(* IEC 61131-3 sources: plcassist-cli/packages/volt-lsp-iec/test-corpus/lenze-mid/Device/Plc Logic/Application/Library Manager/CAA Behaviour Model, 12 files *)

(* ---- VERSIONCONSTANTS.gvl ---- *)
VAR_GLOBAL
	GC_BYVERSION : BYTE := 1;
	GC_BYVERSION_1 : BYTE := 0;
END_VAR

(* ---- IFBCOMMAND.itf ---- *)
INTERFACE IFBCOMMAND
END_INTERFACE

METHOD PRVABORT : BOOL
END_METHOD

METHOD PRVCYCLICACTION : BOOL
END_METHOD

METHOD PRVRESETOUTPUTS : BOOL
END_METHOD

METHOD PRVSTART : BOOL
END_METHOD

(* ---- GETSUPPLIERVERSION.fun ---- *)
FUNCTION GETSUPPLIERVERSION : WORD
VAR_INPUT
	XDUMMY : BOOL;
END_VAR
END_FUNCTION

(* ---- ETRIG.fb ---- *)
FUNCTION_BLOCK ETRIG
VAR_INPUT
	XEXECUTE : BOOL;
END_VAR
VAR_OUTPUT
	XDONE : BOOL;
	XBUSY : BOOL;
	XERROR : BOOL;
END_VAR
VAR
	XPREVIOUSEXECUTE : BOOL;
	XPREVIOUSABORTINPROGRESS : BOOL;
	XABORTINPROGRESS : BOOL;
	IERROR : INT;
END_VAR
END_FUNCTION_BLOCK

METHOD PRVABORT : BOOL
END_METHOD

METHOD PRVCYCLICACTION : BOOL
END_METHOD

METHOD PRVRESETOUTPUTS : BOOL
END_METHOD

METHOD PRVSTART : BOOL
END_METHOD

(* ---- ETRIGA.fb ---- *)
FUNCTION_BLOCK ETRIGA
VAR_INPUT
	XEXECUTE : BOOL;
	XABORT : BOOL;
END_VAR
VAR_OUTPUT
	XDONE : BOOL;
	XBUSY : BOOL;
	XERROR : BOOL;
	XABORTED : BOOL;
END_VAR
VAR
	XPREVIOUSABORTINPROGRESS : BOOL;
	XPREVIOUSEXECUTE : BOOL;
	XABORTINPROGRESS : BOOL;
	IERROR : INT;
END_VAR
END_FUNCTION_BLOCK

METHOD PRVABORT : BOOL
END_METHOD

METHOD PRVCYCLICACTION : BOOL
END_METHOD

METHOD PRVRESETOUTPUTS : BOOL
END_METHOD

METHOD PRVSTART : BOOL
END_METHOD

(* ---- ETRIGTL.fb ---- *)
FUNCTION_BLOCK ETRIGTL
VAR_INPUT
	XEXECUTE : BOOL;
	UDITIMELIMIT : UDINT;
END_VAR
VAR_OUTPUT
	XDONE : BOOL;
	XBUSY : BOOL;
	XERROR : BOOL;
END_VAR
VAR
	XPREVIOUSABORTINPROGRESS : BOOL;
	XPREVIOUSEXECUTE : BOOL;
	XABORTINPROGRESS : BOOL;
	XREPEAT : BOOL;
	TKFBSTART : CAA.TICK;
	TKTIMELIMIT : CAA.TICK;
	IERROR : INT;
END_VAR
END_FUNCTION_BLOCK

METHOD PRVABORT : BOOL
END_METHOD

METHOD PRVCYCLICACTION : BOOL
END_METHOD

METHOD PRVRESETOUTPUTS : BOOL
END_METHOD

METHOD PRVSTART : BOOL
END_METHOD

(* ---- ETRIGTLA.fb ---- *)
FUNCTION_BLOCK ETRIGTLA
VAR_INPUT
	XEXECUTE : BOOL;
	XABORT : BOOL;
	UDITIMELIMIT : UDINT;
END_VAR
VAR_OUTPUT
	XDONE : BOOL;
	XBUSY : BOOL;
	XERROR : BOOL;
	XABORTED : BOOL;
END_VAR
VAR
	XPREVIOUSABORTINPROGRESS : BOOL;
	XPREVIOUSEXECUTE : BOOL;
	XABORTINPROGRESS : BOOL;
	XREPEAT : BOOL;
	TKFBSTART : CAA.TICK;
	TKTIMELIMIT : CAA.TICK;
	IERROR : INT;
END_VAR
END_FUNCTION_BLOCK

METHOD PRVABORT : BOOL
END_METHOD

METHOD PRVCYCLICACTION : BOOL
END_METHOD

METHOD PRVRESETOUTPUTS : BOOL
END_METHOD

METHOD PRVSTART : BOOL
END_METHOD

(* ---- ETRIGTO.fb ---- *)
FUNCTION_BLOCK ETRIGTO
VAR_INPUT
	XEXECUTE : BOOL;
	UDITIMEOUT : UDINT;
END_VAR
VAR_OUTPUT
	XDONE : BOOL;
	XBUSY : BOOL;
	XERROR : BOOL;
END_VAR
VAR
	XPREVIOUSABORTINPROGRESS : BOOL;
	XPREVIOUSEXECUTE : BOOL;
	XABORTINPROGRESS : BOOL;
	TKSTART : CAA.TICK;
	TKTIMEOUT : CAA.TICK;
	IERROR : INT;
END_VAR
END_FUNCTION_BLOCK

METHOD PRVABORT : BOOL
END_METHOD

METHOD PRVCYCLICACTION : BOOL
END_METHOD

METHOD PRVRESETOUTPUTS : BOOL
END_METHOD

METHOD PRVSTART : BOOL
END_METHOD

(* ---- ETRIGTOA.fb ---- *)
FUNCTION_BLOCK ETRIGTOA
VAR_INPUT
	XEXECUTE : BOOL;
	XABORT : BOOL;
	UDITIMEOUT : UDINT;
END_VAR
VAR_OUTPUT
	XDONE : BOOL;
	XBUSY : BOOL;
	XERROR : BOOL;
	XABORTED : BOOL;
END_VAR
VAR
	XPREVIOUSABORTINPROGRESS : BOOL;
	XPREVIOUSEXECUTE : BOOL;
	XABORTINPROGRESS : BOOL;
	TKSTART : CAA.TICK;
	TKTIMEOUT : CAA.TICK;
	IERROR : INT;
END_VAR
END_FUNCTION_BLOCK

METHOD PRVABORT : BOOL
END_METHOD

METHOD PRVCYCLICACTION : BOOL
END_METHOD

METHOD PRVRESETOUTPUTS : BOOL
END_METHOD

METHOD PRVSTART : BOOL
END_METHOD

(* ---- ETRIGTOTL.fb ---- *)
FUNCTION_BLOCK ETRIGTOTL
VAR_INPUT
	XEXECUTE : BOOL;
	UDITIMELIMIT : UDINT;
	UDITIMEOUT : UDINT;
END_VAR
VAR_OUTPUT
	XDONE : BOOL;
	XBUSY : BOOL;
	XERROR : BOOL;
END_VAR
VAR
	XPREVIOUSABORTINPROGRESS : BOOL;
	XPREVIOUSEXECUTE : BOOL;
	XABORTINPROGRESS : BOOL;
	XREPEAT : BOOL;
	TKFBSTART : CAA.TICK;
	TKSTART : CAA.TICK;
	TKTIMELIMIT : CAA.TICK;
	TKTIMEOUT : CAA.TICK;
	IERROR : INT;
END_VAR
END_FUNCTION_BLOCK

METHOD PRVABORT : BOOL
END_METHOD

METHOD PRVCYCLICACTION : BOOL
END_METHOD

METHOD PRVRESETOUTPUTS : BOOL
END_METHOD

METHOD PRVSTART : BOOL
END_METHOD

(* ---- ETRIGTOTLA.fb ---- *)
FUNCTION_BLOCK ETRIGTOTLA
VAR_INPUT
	XEXECUTE : BOOL;
	XABORT : BOOL;
	UDITIMELIMIT : UDINT;
	UDITIMEOUT : UDINT;
END_VAR
VAR_OUTPUT
	XDONE : BOOL;
	XBUSY : BOOL;
	XERROR : BOOL;
	XABORTED : BOOL;
END_VAR
VAR
	XPREVIOUSABORTINPROGRESS : BOOL;
	XPREVIOUSEXECUTE : BOOL;
	XABORTINPROGRESS : BOOL;
	XREPEAT : BOOL;
	TKFBSTART : CAA.TICK;
	TKSTART : CAA.TICK;
	TKTIMELIMIT : CAA.TICK;
	TKTIMEOUT : CAA.TICK;
	IERROR : ERROR;
END_VAR
END_FUNCTION_BLOCK

METHOD PRVABORT : BOOL
END_METHOD

METHOD PRVCYCLICACTION : BOOL
END_METHOD

METHOD PRVRESETOUTPUTS : BOOL
END_METHOD

METHOD PRVSTART : BOOL
END_METHOD

(* ---- LTRIG.fb ---- *)
FUNCTION_BLOCK LTRIG
VAR_INPUT
	XENABLE : BOOL;
END_VAR
VAR_OUTPUT
	XDONE : BOOL;
	XBUSY : BOOL;
	XERROR : BOOL;
END_VAR
VAR
	XPREVIOUSABORTINPROGRESS : BOOL;
	XPREVIOUSENABLE : BOOL;
	XABORTINPROGRESS : BOOL;
	IERROR : INT;
END_VAR
END_FUNCTION_BLOCK

METHOD PRVABORT : BOOL
END_METHOD

METHOD PRVCYCLICACTION : BOOL
END_METHOD

METHOD PRVRESETOUTPUTS : BOOL
END_METHOD

METHOD PRVSTART : BOOL
END_METHOD
